(* IEC 61131-3 sources: codesys-ai-industrial-robot-control/plc/src/Config, 5 files *)

(* ---- GVL_AlarmDefs.st ---- *)
// Alarm definitions: class and operator text for every E_AlarmId.
// Critical -> PackML Abort, Error -> Stop, Warning -> no state change (BinFull suspends the unit).
{attribute 'qualified_only'}
VAR_GLOBAL CONSTANT
    aDefs : ARRAY[E_AlarmId.None..E_AlarmId.QueueOverflow] OF ST_AlarmDef := [
        (eClass := E_AlarmClass.Info, sText := 'No alarm'),
        (eClass := E_AlarmClass.Critical, sText := 'Emergency stop pressed'),
        (eClass := E_AlarmClass.Critical, sText := 'Safety door opened in automatic mode'),
        (eClass := E_AlarmClass.Critical, sText := 'Connection to the digital twin bridge lost'),
        (eClass := E_AlarmClass.Critical, sText := 'Robot axis group error'),
        (eClass := E_AlarmClass.Error, sText := 'Conveyor axis error'),
        (eClass := E_AlarmClass.Warning, sText := 'Joint following error above warning limit'),
        (eClass := E_AlarmClass.Critical, sText := 'Joint following error above fault limit'),
        (eClass := E_AlarmClass.Critical, sText := 'Joint feedback not updated'),
        (eClass := E_AlarmClass.Error, sText := 'Vacuum not reached - part not gripped'),
        (eClass := E_AlarmClass.Error, sText := 'Vacuum lost while carrying a part'),
        (eClass := E_AlarmClass.Warning, sText := 'Part left the pick window unpicked'),
        (eClass := E_AlarmClass.Warning, sText := 'A bin is full - cell suspended until it is emptied'),
        (eClass := E_AlarmClass.Warning, sText := 'No vision result for a captured part'),
        (eClass := E_AlarmClass.Warning, sText := 'AI decision late - fallback rule used'),
        (eClass := E_AlarmClass.Warning, sText := 'Low detection confidence - part quarantined'),
        (eClass := E_AlarmClass.Error, sText := 'Part queue full')];
END_VAR

(* ---- GVL_CellGeometry.st ---- *)
// Fixed geometry of the cell. Units: mm and degrees, robot base frame (Z up).
// Kinematics values must match the axis group AxisGroup_Robot (plc/scripts/build_softmotion_base.py).
// Orientations (A, B, C): B = 180 points the tool straight down (verified in simulation).
{attribute 'qualified_only'}
VAR_GLOBAL CONSTANT
    // Kin_ArticulatedRobot_6DOF parameters [mm]
    ROBOT_A1 : LREAL := 50;
    ROBOT_D1 : LREAL := 400;
    ROBOT_A2 : LREAL := 450;
    ROBOT_A3 : LREAL := 50;
    ROBOT_D3 : LREAL := 0;
    ROBOT_D4 : LREAL := 450;
    ROBOT_D6 : LREAL := 120;                 // flange + suction tool

    // Tool pointing straight down
    TOOL_DOWN_A : LREAL := 0;
    TOOL_DOWN_B : LREAL := 180;
    TOOL_DOWN_C : LREAL := 180;

    // Conveyor belt frame: origin at the infeed, +X along the flow direction.
    BELT_ORIGIN : MC_COORD_REF := (X := -1500, Y := -550, Z := 0, A := 0, B := 0, C := 0);
    BELT_SURFACE_Z : LREAL := 0;
    PE1_X : LREAL := 300;                    // camera trigger photo-eye, belt frame [mm]
    PE2_X : LREAL := 1050;                   // pick window start, belt frame [mm]
    PICK_WINDOW_END_X : LREAL := 1750;       // pick window end, belt frame [mm]
    PICK_MARGIN : LREAL := 300;              // do not start a pick this close to the window end [mm]
    // Grip height of each part class above the belt [mm]: the top surface under the suction
    // cup (config/parts.yaml classes, tools/fetch_objects.py meta.json; a unit test keeps
    // both equal)
    PART_HEIGHTS : ARRAY[0..2] OF LREAL := [56.39, 81.19, 83.46];

    // Home position, joint space [deg]
    HOME_ACS : SMC_POS_REF := (a := (a0 := 0, a1 := -30, a2 := 60, a3 := 0, a4 := 60, a5 := 0));
    // Waiting pose above the pick window, tool down (machine coordinates)
    READY_POSE : MC_COORD_REF := (X := -100, Y := -550, Z := 300, A := 0, B := 180, C := 180);
    RETRACT_HEIGHT : LREAL := 100;           // lift above the bin drop pose after release [mm]

    // Drop poses above the bins (tool pointing down), machine coordinates [mm, deg]. Z 300: a
    // held part up to 90 mm tall clears the 160 mm bin rim by 50 mm.
    BIN_DROP : ARRAY[E_Bin.TypeA..E_Bin.Quarantine] OF MC_COORD_REF := [
        (X := -500, Y := 550, Z := 300, A := 0, B := 180, C := 180),
        (X := -300, Y := 550, Z := 300, A := 0, B := 180, C := 180),
        (X := -100, Y := 550, Z := 300, A := 0, B := 180, C := 180),
        (X := 100, Y := 550, Z := 300, A := 0, B := 180, C := 180),
        (X := 300, Y := 550, Z := 300, A := 0, B := 180, C := 180),
        (X := 500, Y := 550, Z := 300, A := 0, B := 180, C := 180)];
END_VAR

(* ---- GVL_Config.st ---- *)
// Build/run configuration.
{attribute 'qualified_only'}
VAR_GLOBAL
    // Joint feedback := setpoint (no staleness check) unless the twin reports itself active through
    // GVL_Bridge.xTwinActive. FALSE forces real feedback even without the twin.
    xFeedbackLoopback : BOOL := TRUE;
    // The sorting cell runs in PRG_Main. Simulation tests of single blocks switch it off so their
    // harnesses can own the robot and the conveyor.
    xCellEnabled : BOOL := TRUE;
END_VAR
VAR_GLOBAL CONSTANT
    MAX_PARTS : UINT := 32;                  // capacity of the part queue
END_VAR

(* ---- GVL_Constants.st ---- *)
// Project-wide constants. Values that change per recipe live in GVL_Params, not here.
{attribute 'qualified_only'}
VAR_GLOBAL CONSTANT
    PROJECT_VERSION : STRING := '0.7.0';
END_VAR

(* ---- GVL_Params.st ---- *)
// Process parameters. Retained; written by the recipes (Standard / HighSpeed).
{attribute 'qualified_only'}
VAR_GLOBAL RETAIN
    lrBeltSpeed : LREAL := 100;              // conveyor speed [mm/s]
    lrApproachHeight : LREAL := 80;          // approach / lift height above the part [mm]
    lrPickDepth : LREAL := 5;                // how far below the part top the cup goes [mm]
    lrLinVelocity : LREAL := 500;            // linear path velocity [mm/s]
    lrLinAccel : LREAL := 2000;              // linear path acceleration [mm/s2]
    lrLinJerk : LREAL := 20000;              // linear path jerk [mm/s3]
    lrPtpVelFactor : LREAL := 0.5;           // PTP velocity factor ]0, 1]
    rConfidenceThreshold : REAL := 0.6;      // below this the part goes to quarantine
    tDecisionDeadline : TIME := T#2S500MS;   // fallback if no decision by then
    tVacuumTimeout : TIME := T#500MS;        // no grip -> error
    lrFollowErrWarn : LREAL := 2.0;          // following error warning [deg]
    lrFollowErrFault : LREAL := 5.0;         // following error fault [deg]
    tFeedbackTimeout : TIME := T#500MS;      // joint feedback must update within this time
    aClassToBin : ARRAY[0..2] OF E_Bin := [E_Bin.TypeA, E_Bin.TypeB, E_Bin.TypeC];
END_VAR
